Fanuc KAREL source: kc00021.KL

-- PROVISIONAL review KL for V940-1; original PC SHA256 05b54e1dc6da1ecc5ed8a950bcc74e21abca493a99a6bb9d799096157f9d8ca9
-- Incomplete behavior may be omitted. Consult companion uncertainty JSON. Do not deploy.
PROGRAM KC00021
%NOLOCKGROUP
BEGIN
  -- V9_ZERO_TABLE_METADATA_HINT layout=0002_ascii; no indexed target words; source/name/runtime held
  -- UNRESOLVED_PC offsets 5-18; opcodes 27,27,27,9C,31,23
  -- UNRESOLVED_PC offsets 23-27; opcodes 7F
END KC00021
